TYPE "ST_ReleaseReason"
VERSION : 0.1
   STRUCT
      Description : WString[255];
      ReasonCode : DInt;
      SourcePath : WString[255];
      Kind : DInt;
      Bypassable : Bool;
   END_STRUCT;

END_TYPE

